TYPE ST_EL1918_TwinSafe :
STRUCT
	
//EtherCAT Terminal, 8-channel digital input, 
//24 V DC, TwinSAFE, TwinSAFE Logic

	State	AT %I*: UINT;
	i_ch1	AT %I*: BOOL;
	i_ch2	AT %I*: BOOL;
	i_ch3	AT %I*: BOOL;
	i_ch4	AT %I*: BOOL;
	i_ch5	AT %I*: BOOL;
	i_ch6	AT %I*: BOOL;
	i_ch7	AT %I*: BOOL;
	i_ch8	AT %I*: BOOL;
	
END_STRUCT
END_TYPE

(* stored: Version 1.1.0.1, ProductVersion 3.1.4024.12
   DUT ST_EL1918_TwinSafe: Id {d6cf9bd5-66b2-4537-96b2-43cd0f2646ba} *)
